// ---- DUTs/ST_MoverStatus.TcDUT
// C# 端對應 MoverStatus (Pack = 1)
{attribute 'pack_mode' := '1'}
TYPE ST_MoverStatus :
STRUCT
    fPositionMm : LREAL;    // 環上位置 (mm), 0~3000
    fVelocityMmS : LREAL;   // 實際速度 (mm/s)
    bPowered : BOOL;
    bBusy : BOOL;
    bDone : BOOL;
    bError : BOOL;
    nErrorId : UDINT;
    bHasPart : BOOL;        // 有工件
    bPressed : BOOL;        // 已下壓
    nStation : INT;         // 停在哪一站，0 = 不在站上
END_STRUCT
END_TYPE

// ---- DUTs/ST_StationStatus.TcDUT
// C# 端對應 StationStatus (Pack = 1)
{attribute 'pack_mode' := '1'}
TYPE ST_StationStatus :
STRUCT
    eState : E_StationState;
    nStep : INT;            // 站內步驟，見 README
    bOccupied : BOOL;       // 站內有 mover 或站在動作
    nMover : INT;           // 處理中的 mover，0 = 無
    bError : BOOL;
    nErrorId : UDINT;
    nDoneCount : UDINT;     // 完成次數
    fAxis1Mm : LREAL;       // X (mm)；下壓站不用
    fAxis2Mm : LREAL;       // Y (mm)；下壓站不用
    fAxis3Mm : LREAL;       // Z (mm)，往下為正
    bGripClosed : BOOL;     // 夾爪閉合；下壓站固定 FALSE
END_STRUCT
END_TYPE

// ---- GVLs/GVL_ErrorId.TcGVL
// 應用程式錯誤碼；MC / NC 的錯誤碼照原值傳出
{attribute 'qualified_only'}
VAR_GLOBAL CONSTANT
    cErrInvalidState : UDINT := 16#E001;        // 狀態機進到未定義狀態
    cErrMoveTimeout : UDINT := 16#E101;         // mover 移動逾時
    cErrStationTimeout : UDINT := 16#E201;      // 站內步驟逾時
    cErrInitTimeout : UDINT := 16#E301;         // 初始化步驟逾時
    cErrEnvInit : UDINT := 16#E302;             // Utility 環境 Init 失敗
    cErrIdDetection : UDINT := 16#E303;         // Mover ID detection 失敗
    cErrGroup : UDINT := 16#E304;               // CA group enable 失敗
    cErrLostReady : UDINT := 16#E310;           // 執行中掉出可控
    cErrCycle : UDINT := 16#E401;               // 自動循環失敗
END_VAR

// ---- GVLs/GVL_Param.TcGVL
{attribute 'qualified_only'}
VAR_GLOBAL CONSTANT
    cMoverCount : INT := 4;                     // mover 數，與 XTS 設定一致
    cStationCount : INT := 3;                   // 站數
    cStationLoad : INT := 1;                    // 站號：Load
    cStationPress : INT := 2;                   // 站號：Press
    cStationUnload : INT := 3;                  // 站號：Unload
    cTrackLengthMm : LREAL := 3000.0;           // 軌道長 (mm)
    cStationPosMm : ARRAY[1..3] OF LREAL := [1600.0, 2100.0, 2600.0];   // 各站 mover 停止位置 (mm, 環上)
    cMaxVelocityMmS : LREAL := 1500.0;          // mover 速度上限 (mm/s)
    cDefaultVelocityMmS : LREAL := 400.0;       // 自動循環 / 送站速度 (mm/s)
    cMoverAccMmS2 : LREAL := 2000.0;            // mover 加減速度 (mm/s2)
    cMoverJerkMmS3 : LREAL := 20000.0;          // mover jerk (mm/s3)
    cCaGapMm : LREAL := 110.0;                  // CA 最小間距 (mm)
    cAtStationTolMm : LREAL := 1.0;             // 判定到站的容差 (mm)
    cMoveTimeout : TIME := T#10M;               // mover 單次移動上限
    cInitStepTimeout : TIME := T#5M;            // 初始化每一步上限，UmRT 偏慢所以放寬
    cResetTime : TIME := T#500MS;               // 初始化 reset 保持時間
    cStationStepTimeout : TIME := T#2M;         // 站內每一步上限
    cGantryAxisCount : INT := 3;                // XYZ 軸數
    cAxisX : INT := 1;
    cAxisY : INT := 2;
    cAxisZ : INT := 3;
    cGantryVelocityMmS : LREAL := 200.0;        // XYZ 與下壓軸速度 (mm/s)
    cGantryAccMmS2 : LREAL := 1000.0;           // XYZ 與下壓軸加減速度 (mm/s2)
    cGantryZUpMm : LREAL := 0.0;                // Z 上位 (mm)
    cGantryZDownMm : LREAL := 80.0;             // Z 下位 (mm)
    cGantryFeederXMm : LREAL := 300.0;          // Load 取料點 X (mm)
    cGantryFeederYMm : LREAL := 150.0;          // Load 取料點 Y (mm)
    cGantryOutXMm : LREAL := 300.0;             // Unload 放料點 X (mm)
    cGantryOutYMm : LREAL := -150.0;            // Unload 放料點 Y (mm)
    cGantryMoverXMm : LREAL := 0.0;             // mover 正上方 X (mm)
    cGantryMoverYMm : LREAL := 0.0;             // mover 正上方 Y (mm)
    cGripTime : TIME := T#300MS;                // 夾 / 放 時間
    cPressZDownMm : LREAL := 50.0;              // 下壓位置 (mm)
    cPressHoldTime : TIME := T#1S;              // 保壓時間
END_VAR

// ---- POUs/MAIN.TcPOU
PROGRAM MAIN
VAR
    aAxis : ARRAY[1..GVL_Param.cMoverCount] OF AXIS_REF;              // 連 NC Mover Axis 1..4
    stCaGroup : Tc3_McCoordinatedMotion.AXES_GROUP_REF;                 // 連 XtsCaGroup
    aLoadAxis : ARRAY[1..GVL_Param.cGantryAxisCount] OF AXIS_REF;      // 連 Load X / Y / Z
    aUnloadAxis : ARRAY[1..GVL_Param.cGantryAxisCount] OF AXIS_REF;    // 連 Unload X / Y / Z
    stPressAxis : AXIS_REF;                                             // 連 Press Z
    fbXts : FB_XTS_Control;                                             // C# RPC 主入口：MAIN.fbXts
    refMover1 : REFERENCE TO FB_Mover;                                  // 備案 RPC 路徑：MAIN.refMover1..4
    refMover2 : REFERENCE TO FB_Mover;
    refMover3 : REFERENCE TO FB_Mover;
    refMover4 : REFERENCE TO FB_Mover;
END_VAR

fbXts(aMoverAxis := aAxis, stGroup := stCaGroup, aLoadAxis := aLoadAxis,
    aUnloadAxis := aUnloadAxis, stPressAxis := stPressAxis);
// REFERENCE 每 cycle 重取 (PTR-03)
refMover1 REF= fbXts.M_GetMover(1);
refMover2 REF= fbXts.M_GetMover(2);
refMover3 REF= fbXts.M_GetMover(3);
refMover4 REF= fbXts.M_GetMover(4);

END_PROGRAM

// ---- POUs/FB_XTS_Control.TcPOU
// 整線總控：初始化 (Find mover 1 → 送電 → CA group)、模式、自動循環 Load → Press → Unload、派 mover 到站。
// 擁有 4 個 FB_Mover 與 3 個站；每 cycle 把 ST_CmdPermit 寫給子 FB，所有命令檢查只走 F_CheckCmdAllowed。
FUNCTION_BLOCK FB_XTS_Control
VAR_IN_OUT
    aMoverAxis : ARRAY[1..GVL_Param.cMoverCount] OF AXIS_REF;          // XTS mover NC 軸
    stGroup : Tc3_McCoordinatedMotion.AXES_GROUP_REF;                   // CA group
    aLoadAxis : ARRAY[1..GVL_Param.cGantryAxisCount] OF AXIS_REF;      // Load 站 XYZ
    aUnloadAxis : ARRAY[1..GVL_Param.cGantryAxisCount] OF AXIS_REF;    // Unload 站 XYZ
    stPressAxis : AXIS_REF;                                             // Press 站下壓軸
END_VAR
VAR_OUTPUT
    bReady : BOOL;                  // 可控
    eMode : E_XtsMode;
    eInitStep : E_InitStep;
    eCycleState : E_CycleState;
    bError : BOOL;
    nErrorId : UDINT;
END_VAR
VAR
    aMover : ARRAY[1..GVL_Param.cMoverCount] OF FB_Mover;
    fbLoad : FB_StationLoad;
    fbPress : FB_StationPress;
    fbUnload : FB_StationUnload;
    aStationPtr : ARRAY[1..GVL_Param.cStationCount] OF POINTER TO FB_Station;   // 每 cycle 重取
    fbEnvironment : Tc3_XTS_Utility.FB_TcIoXtsEnvironment;
    stEnvConfig : Tc3_XTS_Utility.ST_XtsEnvironmentConfiguration;
    fbGroup : FB_CaGroup;
    fbInitTimer : TON;
    fbResetTimer : TON;
    stPermit : ST_CmdPermit;
    stStatus : ST_LineStatus;       // M_GetStatus 回傳的快照
    sInitMsg : STRING;              // 初始化進度或失敗原因
    sCycleMsg : STRING;             // 自動循環訊息
    bEnvInitialized : BOOL;
    bPowerOn : BOOL;
    bGroupEnable : BOOL;
    bInitReset : BOOL;
    eInitStepLast : E_InitStep;
    tInitStart : TIME;              // M_InitialXTS 被取走的時刻
    nFindMover1Ms : UDINT;          // 各步完成時間 (ms，從 tInitStart 起算；0 = 這次還沒完成)
    bFindMover1Detected : BOOL;     // TRUE = detection valid；FALSE 且 nFindMover1Ms > 0 = 跳過
    nPowerOnMs : UDINT;
    nGroupMs : UDINT;
    bReqInit : BOOL;                // method 設，body 取走
    bReqStop : BOOL;
    bReqSetMode : BOOL;
    eReqMode : E_XtsMode;
    bReqStartCycle : BOOL;
    nReqCycleMover : INT;
    bStopPulse : BOOL;              // 本 cycle 對站送 abort
    nCycleMover : INT;
    nCycleStation : INT;
    bCycleMoveIssued : BOOL;
    nCycleCount : UDINT;
    tCycleStart : TIME;
    aStationDoneMs : ARRAY[1..GVL_Param.cStationCount] OF UDINT;
    aLastDoneCount : ARRAY[1..GVL_Param.cStationCount] OF UDINT;
    aMoverAtStation : ARRAY[1..GVL_Param.cStationCount] OF INT;
    pStation : POINTER TO FB_Station;
    bAllPowered : BOOL;
    bAnyMoverError : BOOL;
    bInitBusy : BOOL;
    fDistMm : LREAL;
    i : INT;
    j : INT;
    nStation : INT;
END_VAR

// 1. 站指標每 cycle 重取 (PTR-03)
aStationPtr[GVL_Param.cStationLoad] := ADR(fbLoad);
aStationPtr[GVL_Param.cStationPress] := ADR(fbPress);
aStationPtr[GVL_Param.cStationUnload] := ADR(fbUnload);

// 2. 取走 method 設的命令
bStopPulse := FALSE;
IF bReqStop THEN
    bReqStop := FALSE;
    bStopPulse := TRUE;
    FOR i := 1 TO GVL_Param.cMoverCount DO
        aMover[i].M_Stop();
    END_FOR
    IF (eCycleState = E_CycleState.ToStation) OR (eCycleState = E_CycleState.InStation) THEN
        eCycleState := E_CycleState.Stopped;
        sCycleMsg := 'Stopped by M_Stop';
    END_IF
END_IF
IF bReqSetMode THEN
    bReqSetMode := FALSE;
    eMode := eReqMode;
END_IF
IF bReqInit THEN
    bReqInit := FALSE;
    bError := FALSE;
    nErrorId := 0;
    sInitMsg := 'Reset';
    eInitStep := E_InitStep.Reset;
    tInitStart := TIME();
    nFindMover1Ms := 0;
    bFindMover1Detected := FALSE;
    nPowerOnMs := 0;
    nGroupMs := 0;
END_IF

// 3. 初始化：Find mover 1 → 送電 → CA group
bInitBusy := M_InitBusy();
fbInitTimer(IN := bInitBusy AND (eInitStep = eInitStepLast), PT := GVL_Param.cInitStepTimeout);
eInitStepLast := eInitStep;
fbResetTimer(IN := (eInitStep = E_InitStep.Reset), PT := GVL_Param.cResetTime);
CASE eInitStep OF
E_InitStep.Idle, E_InitStep.Ready, E_InitStep.Error:
    ;
E_InitStep.Reset:
    bInitReset := TRUE;
    bPowerOn := FALSE;
    bGroupEnable := FALSE;
    IF fbResetTimer.Q THEN
        bInitReset := FALSE;
        IF bEnvInitialized THEN
            eInitStep := E_InitStep.WaitMovers;
        ELSE
            stEnvConfig.bEnableInitInfoServer := TRUE;
            stEnvConfig.bEnableInitCaGroup := TRUE;
            fbEnvironment.P_XtsEnvironmentConfiguration := stEnvConfig;
            eInitStep := E_InitStep.InitEnvironment;
        END_IF
        sInitMsg := F_InitStepName(eInitStep);
    END_IF
E_InitStep.InitEnvironment:
    // Init 是非同步的，回 TRUE 才算做完
    IF fbEnvironment.Init(TRUE) THEN
        fbEnvironment.Init(FALSE);
        IF fbEnvironment.P_IsInitialized THEN
            bEnvInitialized := TRUE;
            eInitStep := E_InitStep.WaitMovers;
            sInitMsg := F_InitStepName(eInitStep);
        ELSE
            M_SetInitError(nId := GVL_ErrorId.cErrEnvInit, sText := 'Tc3_XTS_Utility Init failed');
        END_IF
    END_IF
E_InitStep.WaitMovers:
    IF (fbEnvironment.XpuTcIo(1).GetDetectedMoverCount() = INT_TO_UDINT(GVL_Param.cMoverCount))
        AND fbEnvironment.XpuTcIo(1).GetAreAllPositionsValid() THEN
        eInitStep := E_InitStep.FindMover1;
        sInitMsg := F_InitStepName(eInitStep);
    END_IF
E_InitStep.FindMover1:
    // 專案設定 IdDetectionMode = Mover1；detection 要在 MC_Power 之前 (XTS 事件 9016)
    IF fbEnvironment.XpuTcIo(1).GetMoverIdDetectionMode() = MoverIdDetectionMode.Mover1 THEN
        IF fbEnvironment.XpuTcIo(1).TriggerMoverIdDetection() THEN
            eInitStep := E_InitStep.FindMover1Wait;
            sInitMsg := 'FindMover1: Mover ID detection triggered, waiting for result';
        ELSE
            M_SetInitError(nId := GVL_ErrorId.cErrIdDetection, sText := 'TriggerMoverIdDetection rejected');
        END_IF
    ELSE
        // 防呆：XPU 被改回 Standard 時不做 detection，mover 編號照設定順序
        eInitStep := E_InitStep.PowerOn;
        sInitMsg := 'FindMover1 skipped: XPU IdDetectionMode is not Mover1, PowerOn';
        nFindMover1Ms := MAX(TIME_TO_UDINT(TIME() - tInitStart), 1);
    END_IF
E_InitStep.FindMover1Wait:
    IF fbEnvironment.XpuTcIo(1).GetHasMoverIdDetectionError() THEN
        M_SetInitError(nId := GVL_ErrorId.cErrIdDetection, sText := 'Mover ID detection error');
    ELSIF fbEnvironment.XpuTcIo(1).GetIsMoverIdDetectionValid() THEN
        eInitStep := E_InitStep.PowerOn;
        sInitMsg := 'FindMover1 done (Mover ID detection valid), PowerOn';
        nFindMover1Ms := MAX(TIME_TO_UDINT(TIME() - tInitStart), 1);
        bFindMover1Detected := TRUE;
    END_IF
E_InitStep.PowerOn:
    bPowerOn := TRUE;
    IF bAllPowered AND fbLoad.bAxesPowered AND fbPress.bAxesPowered AND fbUnload.bAxesPowered THEN
        eInitStep := E_InitStep.EnableGroup;
        sInitMsg := F_InitStepName(eInitStep);
        nPowerOnMs := MAX(TIME_TO_UDINT(TIME() - tInitStart), 1);
    END_IF
E_InitStep.EnableGroup:
    bGroupEnable := TRUE;
    IF fbGroup.bError THEN
        M_SetInitError(nId := fbGroup.nErrorId, sText := 'CA group error');
    ELSIF fbGroup.bReady THEN
        eInitStep := E_InitStep.Ready;
        sInitMsg := 'Ready';
        nGroupMs := MAX(TIME_TO_UDINT(TIME() - tInitStart), 1);
    END_IF
ELSE
    M_SetInitError(nId := GVL_ErrorId.cErrInvalidState, sText := 'invalid init step');
END_CASE
IF fbInitTimer.Q THEN
    M_SetInitError(nId := GVL_ErrorId.cErrInitTimeout, sText := 'step timeout');
END_IF

// 4. 可控監視：任何 mover error、失電、group 失效、站上軸 error 都掉出 ready
bAllPowered := TRUE;
bAnyMoverError := FALSE;
FOR i := 1 TO GVL_Param.cMoverCount DO
    bAllPowered := bAllPowered AND aMover[i].bPowered;
    bAnyMoverError := bAnyMoverError OR aMover[i].bError;
END_FOR
IF eInitStep = E_InitStep.Ready THEN
    IF bAnyMoverError THEN
        M_SetInitError(nId := GVL_ErrorId.cErrLostReady, sText := 'mover error');
    ELSIF NOT bAllPowered THEN
        M_SetInitError(nId := GVL_ErrorId.cErrLostReady, sText := 'mover power lost');
    ELSIF NOT fbGroup.bReady THEN
        M_SetInitError(nId := GVL_ErrorId.cErrLostReady, sText := 'CA group not ready');
    ELSIF fbLoad.bAxisError OR fbPress.bAxisError OR fbUnload.bAxisError THEN
        M_SetInitError(nId := GVL_ErrorId.cErrLostReady, sText := 'station axis error');
    END_IF
END_IF
bReady := (eInitStep = E_InitStep.Ready);
stPermit.bReady := bReady;
stPermit.eMode := eMode;

// 5. 哪個 mover 停在哪一站 (停止且在容差內)
FOR nStation := 1 TO GVL_Param.cStationCount DO
    aMoverAtStation[nStation] := 0;
    FOR i := 1 TO GVL_Param.cMoverCount DO
        fDistMm := F_RingPosition(fPositionMm := aMover[i].fPositionMm - GVL_Param.cStationPosMm[nStation]
            + GVL_Param.cTrackLengthMm / 2.0, fLengthMm := GVL_Param.cTrackLengthMm) - GVL_Param.cTrackLengthMm / 2.0;
        IF NOT aMover[i].bBusy AND (ABS(fDistMm) <= GVL_Param.cAtStationTolMm) THEN
            aMoverAtStation[nStation] := i;
        END_IF
    END_FOR
    pStation := aStationPtr[nStation];
    IF pStation <> 0 THEN
        pStation^.nMoverAtStation := aMoverAtStation[nStation];
        j := aMoverAtStation[nStation];
        IF j > 0 THEN
            pStation^.bMoverHasPart := aMover[j].bHasPart;
            pStation^.bMoverPressed := aMover[j].bPressed;
        ELSE
            pStation^.bMoverHasPart := FALSE;
            pStation^.bMoverPressed := FALSE;
        END_IF
    END_IF
END_FOR

// 6. 站完成 → 更新 mover 工件狀態 (手動與自動都走這裡)
FOR nStation := 1 TO GVL_Param.cStationCount DO
    pStation := aStationPtr[nStation];
    IF pStation <> 0 THEN
        IF pStation^.nDoneCount <> aLastDoneCount[nStation] THEN
            aLastDoneCount[nStation] := pStation^.nDoneCount;
            j := pStation^.nMover;
            IF (j >= 1) AND (j <= GVL_Param.cMoverCount) THEN
                CASE nStation OF
                GVL_Param.cStationLoad:
                    aMover[j].M_SetPart(bPart := TRUE, bPress := FALSE);
                GVL_Param.cStationPress:
                    aMover[j].M_SetPart(bPart := aMover[j].bHasPart, bPress := TRUE);
                GVL_Param.cStationUnload:
                    aMover[j].M_SetPart(bPart := FALSE, bPress := FALSE);
                END_CASE
            END_IF
        END_IF
    END_IF
END_FOR

// 7. 自動循環：mover 依序到 Load → Press → Unload
IF NOT bReady AND ((eCycleState = E_CycleState.ToStation) OR (eCycleState = E_CycleState.InStation)) THEN
    eCycleState := E_CycleState.Error;
    sCycleMsg := 'Lost ready during cycle';
END_IF
pStation := 0;
IF (nCycleStation >= 1) AND (nCycleStation <= GVL_Param.cStationCount) THEN
    pStation := aStationPtr[nCycleStation];
END_IF
CASE eCycleState OF
E_CycleState.Idle, E_CycleState.Done, E_CycleState.Stopped, E_CycleState.Error:
    IF bReqStartCycle THEN
        nCycleMover := nReqCycleMover;
        nCycleStation := GVL_Param.cStationLoad;
        bCycleMoveIssued := FALSE;
        tCycleStart := TIME();
        FOR nStation := 1 TO GVL_Param.cStationCount DO
            aStationDoneMs[nStation] := 0;
        END_FOR
        sCycleMsg := 'Cycle started';
        eCycleState := E_CycleState.ToStation;
    END_IF
E_CycleState.ToStation:
    IF pStation = 0 THEN
        eCycleState := E_CycleState.Error;
        sCycleMsg := 'Invalid station index';
    ELSIF NOT bCycleMoveIssued THEN
        bCycleMoveIssued := aMover[nCycleMover].M_RequestMove(fPosition := GVL_Param.cStationPosMm[nCycleStation],
            fVelocity := GVL_Param.cDefaultVelocityMmS, sMsg => sCycleMsg);
    ELSIF aMover[nCycleMover].bDone AND (aMoverAtStation[nCycleStation] = nCycleMover) THEN
        IF pStation^.M_RequestStart(sMsg => sCycleMsg) THEN
            eCycleState := E_CycleState.InStation;
        ELSE
            eCycleState := E_CycleState.Error;
        END_IF
    END_IF
E_CycleState.InStation:
    IF pStation = 0 THEN
        eCycleState := E_CycleState.Error;
        sCycleMsg := 'Invalid station index';
    ELSIF pStation^.eState = E_StationState.Error THEN
        eCycleState := E_CycleState.Error;
        sCycleMsg := 'Station error';
    ELSIF pStation^.eState = E_StationState.Done THEN
        aStationDoneMs[nCycleStation] := TIME_TO_UDINT(TIME() - tCycleStart);
        pStation^.M_RequestRelease(sMsg => sCycleMsg);
        IF nCycleStation < GVL_Param.cStationCount THEN
            nCycleStation := nCycleStation + 1;
            bCycleMoveIssued := FALSE;
            eCycleState := E_CycleState.ToStation;
        ELSE
            nCycleCount := nCycleCount + 1;
            sCycleMsg := 'Cycle done';
            eCycleState := E_CycleState.Done;
        END_IF
    END_IF
ELSE
    eCycleState := E_CycleState.Error;
    sCycleMsg := 'Invalid cycle state';
END_CASE
bReqStartCycle := FALSE;

// 8. 呼叫子 FB (每 cycle 無條件)
FOR i := 1 TO GVL_Param.cMoverCount DO
    aMover[i](nIndex := i, stPermit := stPermit, bPowerEnable := bPowerOn, bResetCmd := bInitReset,
        stAxis := aMoverAxis[i]);
END_FOR
fbGroup(Group := stGroup, Axes := aMoverAxis, bEnable := bGroupEnable, bReset := bInitReset);
fbLoad(nIndex := GVL_Param.cStationLoad, stPermit := stPermit, bPowerEnable := bPowerOn,
    bResetCmd := bInitReset, bAbort := bStopPulse, aAxis := aLoadAxis);
fbPress(nIndex := GVL_Param.cStationPress, stPermit := stPermit, bPowerEnable := bPowerOn,
    bResetCmd := bInitReset, bAbort := bStopPulse, stAxis := stPressAxis);
fbUnload(nIndex := GVL_Param.cStationUnload, stPermit := stPermit, bPowerEnable := bPowerOn,
    bResetCmd := bInitReset, bAbort := bStopPulse, aAxis := aUnloadAxis);

// 9. 狀態快照
stStatus.bReady := bReady;
stStatus.eMode := eMode;
stStatus.eInitStep := eInitStep;
stStatus.bError := bError;
stStatus.nErrorId := nErrorId;
stStatus.eCycleState := eCycleState;
stStatus.nCycleMover := nCycleMover;
stStatus.nCycleStation := nCycleStation;
stStatus.nCycleCount := nCycleCount;
FOR i := 1 TO GVL_Param.cMoverCount DO
    stStatus.aMover[i].fPositionMm := aMover[i].fPositionMm;
    stStatus.aMover[i].fVelocityMmS := aMover[i].fVelocityMmS;
    stStatus.aMover[i].bPowered := aMover[i].bPowered;
    stStatus.aMover[i].bBusy := aMover[i].bBusy;
    stStatus.aMover[i].bDone := aMover[i].bDone;
    stStatus.aMover[i].bError := aMover[i].bError;
    stStatus.aMover[i].nErrorId := aMover[i].nErrorId;
    stStatus.aMover[i].bHasPart := aMover[i].bHasPart;
    stStatus.aMover[i].bPressed := aMover[i].bPressed;
    stStatus.aMover[i].nStation := 0;
END_FOR
FOR nStation := 1 TO GVL_Param.cStationCount DO
    stStatus.aStationDoneMs[nStation] := aStationDoneMs[nStation];
    j := aMoverAtStation[nStation];
    IF (j >= 1) AND (j <= GVL_Param.cMoverCount) THEN
        stStatus.aMover[j].nStation := nStation;
    END_IF
    pStation := aStationPtr[nStation];
    IF pStation <> 0 THEN
        stStatus.aStation[nStation] := pStation^.M_GetStatusStruct();
    END_IF
END_FOR

// 內部用：給 MAIN 的 REFERENCE 備案路徑。超出範圍回 mover 1。
METHOD PUBLIC M_GetMover : REFERENCE TO FB_Mover
VAR_INPUT
    nMover : INT;
END_VAR
M_GetMover REF= aMover[LIMIT(1, nMover, GVL_Param.cMoverCount)];
END_METHOD

// RPC：整線快照 (mover、站、XYZ / 下壓軸位置、循環)，隨時可讀
{attribute 'TcRpcEnable'}
METHOD PUBLIC M_GetStatus : BOOL
VAR_OUTPUT
    stLine : ST_LineStatus;
    sCycle : STRING;            // 自動循環訊息
END_VAR
stLine := stStatus;
sCycle := sCycleMsg;
M_GetStatus := TRUE;
END_METHOD

METHOD PRIVATE M_InitBusy : BOOL
M_InitBusy := (eInitStep = E_InitStep.Reset) OR (eInitStep = E_InitStep.InitEnvironment)
    OR (eInitStep = E_InitStep.WaitMovers) OR (eInitStep = E_InitStep.FindMover1)
    OR (eInitStep = E_InitStep.FindMover1Wait) OR (eInitStep = E_InitStep.PowerOn)
    OR (eInitStep = E_InitStep.EnableGroup);
END_METHOD

// RPC：開始初始化 (Reset → Find mover 1 → PowerOn → EnableGroup)。回 TRUE = 已接受，用 M_ReadXTS_Status 看進度。
{attribute 'TcRpcEnable'}
METHOD PUBLIC M_InitialXTS : BOOL
VAR_OUTPUT
    sMsg : STRING;
END_VAR
M_InitialXTS := FALSE;
IF bReqInit THEN
    sMsg := 'Previous command not yet taken by PLC, retry';
ELSIF M_InitBusy() THEN
    sMsg := CONCAT('Init already running: ', F_InitStepName(eInitStep));
ELSIF (eCycleState = E_CycleState.ToStation) OR (eCycleState = E_CycleState.InStation) THEN
    sMsg := 'Cycle running, call M_Stop first';
ELSIF bReady THEN
    sMsg := 'Already ready';
ELSE
    bReqInit := TRUE;
    sMsg := 'Init started';
    M_InitialXTS := TRUE;
END_IF
END_METHOD

// RPC：總控層的 mover 移動 (陣列元素路徑不能用時的備案)。需 ready + Manual。
{attribute 'TcRpcEnable'}
METHOD PUBLIC M_MoveTo : BOOL
VAR_INPUT
    nMover : UINT;              // 1..cMoverCount
    fPosition : LREAL;          // 目標環上位置 (mm)
    fVelocity : LREAL;          // 速度 (mm/s)
END_VAR
VAR_OUTPUT
    sMsg : STRING;
END_VAR
M_MoveTo := FALSE;
IF NOT F_CheckCmdAllowed(stPermit := stPermit, bNeedManual := TRUE, bNeedAuto := FALSE, sMsg => sMsg) THEN
    RETURN;
END_IF
IF (nMover < 1) OR (nMover > INT_TO_UINT(GVL_Param.cMoverCount)) THEN
    sMsg := CONCAT('nMover out of range 1..', INT_TO_STRING(GVL_Param.cMoverCount));
    RETURN;
END_IF
M_MoveTo := aMover[UINT_TO_INT(nMover)].M_RequestMove(fPosition := fPosition, fVelocity := fVelocity, sMsg => sMsg);
END_METHOD

// RPC：可控閘門狀態，隨時可讀
{attribute 'TcRpcEnable'}
METHOD PUBLIC M_ReadXTS_Status : BOOL
VAR_OUTPUT
    bIsReady : BOOL;            // TRUE 才能下站與 mover 命令
    eStep : E_InitStep;         // 初始化目前步驟
    sStepMsg : STRING;          // 進度或失敗原因
    bIsError : BOOL;
    nErrId : UDINT;
    eModeNow : E_XtsMode;
    nFindMover1DoneMs : UDINT;  // 各步完成時間 (PLC ms，從 M_InitialXTS 被取走起算；0 = 這次還沒完成)
    bFindMover1Valid : BOOL;    // TRUE = Mover ID detection valid；FALSE 且時間 > 0 = IdDetectionMode 不是 Mover1、跳過
    nPowerOnDoneMs : UDINT;
    nGroupDoneMs : UDINT;
END_VAR
bIsReady := bReady;
eStep := eInitStep;
sStepMsg := sInitMsg;
bIsError := bError;
nErrId := nErrorId;
eModeNow := eMode;
nFindMover1DoneMs := nFindMover1Ms;
bFindMover1Valid := bFindMover1Detected;
nPowerOnDoneMs := nPowerOnMs;
nGroupDoneMs := nGroupMs;
M_ReadXTS_Status := TRUE;
END_METHOD

// RPC：總控層的手動放行 (備案路徑)。需 ready + Manual。
{attribute 'TcRpcEnable'}
METHOD PUBLIC M_ReleaseStation : BOOL
VAR_INPUT
    nStation : UINT;            // 1 = Load, 2 = Press, 3 = Unload
END_VAR
VAR_OUTPUT
    sMsg : STRING;
END_VAR
VAR
    pSt : POINTER TO FB_Station;
END_VAR
M_ReleaseStation := FALSE;
IF NOT F_CheckCmdAllowed(stPermit := stPermit, bNeedManual := TRUE, bNeedAuto := FALSE, sMsg => sMsg) THEN
    RETURN;
END_IF
IF (nStation < 1) OR (nStation > INT_TO_UINT(GVL_Param.cStationCount)) THEN
    sMsg := CONCAT('nStation out of range 1..', INT_TO_STRING(GVL_Param.cStationCount));
    RETURN;
END_IF
pSt := aStationPtr[UINT_TO_INT(nStation)];
IF pSt = 0 THEN
    sMsg := 'Station not ready yet, retry';
    RETURN;
END_IF
M_ReleaseStation := pSt^.M_RequestRelease(sMsg => sMsg);
END_METHOD

// RPC：把 mover 送到指定站。需 ready + Manual、站號有效、站沒被其他 mover 佔用。
{attribute 'TcRpcEnable'}
METHOD PUBLIC M_SendToStation : BOOL
VAR_INPUT
    nMover : UINT;              // 1..cMoverCount
    nStation : UINT;            // 1 = Load, 2 = Press, 3 = Unload
END_VAR
VAR_OUTPUT
    sMsg : STRING;
END_VAR
VAR
    nMv : INT;
    nSt : INT;
END_VAR
M_SendToStation := FALSE;
IF NOT F_CheckCmdAllowed(stPermit := stPermit, bNeedManual := TRUE, bNeedAuto := FALSE, sMsg => sMsg) THEN
    RETURN;
END_IF
IF (nMover < 1) OR (nMover > INT_TO_UINT(GVL_Param.cMoverCount)) THEN
    sMsg := CONCAT('nMover out of range 1..', INT_TO_STRING(GVL_Param.cMoverCount));
    RETURN;
END_IF
IF (nStation < 1) OR (nStation > INT_TO_UINT(GVL_Param.cStationCount)) THEN
    sMsg := CONCAT('nStation out of range 1..', INT_TO_STRING(GVL_Param.cStationCount));
    RETURN;
END_IF
nMv := UINT_TO_INT(nMover);       // 已檢查範圍，不會溢位
nSt := UINT_TO_INT(nStation);
IF (aMoverAtStation[nSt] <> 0) AND (aMoverAtStation[nSt] <> nMv) THEN
    sMsg := CONCAT(CONCAT('Station occupied by mover ', INT_TO_STRING(aMoverAtStation[nSt])), ', move it away first');
    RETURN;
END_IF
M_SendToStation := aMover[nMv].M_RequestMove(fPosition := GVL_Param.cStationPosMm[nSt],
    fVelocity := GVL_Param.cDefaultVelocityMmS, sMsg => sMsg);
END_METHOD

METHOD PRIVATE M_SetInitError
VAR_INPUT
    nId : UDINT;
    sText : STRING;
END_VAR
sInitMsg := CONCAT(CONCAT(F_InitStepName(eInitStep), ': '), sText);
bError := TRUE;
nErrorId := nId;
IF nErrorId = 0 THEN
    nErrorId := GVL_ErrorId.cErrInvalidState;
END_IF
eInitStep := E_InitStep.Error;
END_METHOD

// RPC：切換模式 0 = Manual、1 = Auto。自動循環中拒絕。不受 ready 限制。
{attribute 'TcRpcEnable'}
METHOD PUBLIC M_SetMode : BOOL
VAR_INPUT
    nMode : INT;                // 0 = Manual, 1 = Auto
END_VAR
VAR_OUTPUT
    sMsg : STRING;
END_VAR
M_SetMode := FALSE;
IF (eCycleState = E_CycleState.ToStation) OR (eCycleState = E_CycleState.InStation) THEN
    sMsg := 'Cycle running, call M_Stop first';
ELSIF nMode = 0 THEN
    eReqMode := E_XtsMode.Manual;
    bReqSetMode := TRUE;
    sMsg := 'Mode -> Manual';
    M_SetMode := TRUE;
ELSIF nMode = 1 THEN
    eReqMode := E_XtsMode.Auto;
    bReqSetMode := TRUE;
    sMsg := 'Mode -> Auto';
    M_SetMode := TRUE;
ELSE
    sMsg := 'nMode must be 0 (Manual) or 1 (Auto)';
END_IF
END_METHOD

// RPC：nMover 跑一輪 Load → Press → Unload。需 ready + Auto、三站 Idle、mover 沒工件、路徑上沒有其他 mover。
{attribute 'TcRpcEnable'}
METHOD PUBLIC M_StartCycle : BOOL
VAR_INPUT
    nMover : UINT;              // 1..cMoverCount
END_VAR
VAR_OUTPUT
    sMsg : STRING;
END_VAR
VAR
    nMv : INT;
    nOther : INT;
    fPathMm : LREAL;            // 到 Unload 的路徑長 + CA 間距 (mm)
    fAheadMm : LREAL;           // 其他 mover 在前方多遠 (mm)
END_VAR
M_StartCycle := FALSE;
IF NOT F_CheckCmdAllowed(stPermit := stPermit, bNeedManual := FALSE, bNeedAuto := TRUE, sMsg => sMsg) THEN
    RETURN;
END_IF
IF bReqStartCycle THEN
    sMsg := 'Previous command not yet taken by PLC, retry';
    RETURN;
END_IF
IF (eCycleState = E_CycleState.ToStation) OR (eCycleState = E_CycleState.InStation) THEN
    sMsg := 'Cycle already running';
    RETURN;
END_IF
IF (nMover < 1) OR (nMover > INT_TO_UINT(GVL_Param.cMoverCount)) THEN
    sMsg := CONCAT('nMover out of range 1..', INT_TO_STRING(GVL_Param.cMoverCount));
    RETURN;
END_IF
nMv := UINT_TO_INT(nMover);       // 已檢查範圍，不會溢位
IF aMover[nMv].bHasPart THEN
    sMsg := 'Mover already has a part, unload it first';
    RETURN;
END_IF
IF aMover[nMv].bBusy OR aMover[nMv].bError THEN
    sMsg := 'Mover busy or in error';
    RETURN;
END_IF
IF (fbLoad.eState <> E_StationState.Idle) OR (fbPress.eState <> E_StationState.Idle)
    OR (fbUnload.eState <> E_StationState.Idle) THEN
    sMsg := 'All stations must be Idle';
    RETURN;
END_IF
// CA 會讓 mover 排在前車後面，路徑上有車就到不了站
fPathMm := F_RingPosition(fPositionMm := GVL_Param.cStationPosMm[GVL_Param.cStationUnload] - aMover[nMv].fPositionMm,
    fLengthMm := GVL_Param.cTrackLengthMm) + GVL_Param.cCaGapMm;
FOR nOther := 1 TO GVL_Param.cMoverCount DO
    IF nOther <> nMv THEN
        fAheadMm := F_RingPosition(fPositionMm := aMover[nOther].fPositionMm - aMover[nMv].fPositionMm,
            fLengthMm := GVL_Param.cTrackLengthMm);
        IF fAheadMm < fPathMm THEN
            sMsg := CONCAT(CONCAT('Mover ', INT_TO_STRING(nOther)), ' is in the path, move it away in Manual first');
            RETURN;
        END_IF
    END_IF
END_FOR
nReqCycleMover := nMv;
bReqStartCycle := TRUE;
sMsg := 'Cycle accepted';
M_StartCycle := TRUE;
END_METHOD

// RPC：總控層的手動站啟動 (子類別上繼承來的 RPC 不能用時的備案)。需 ready + Manual。
{attribute 'TcRpcEnable'}
METHOD PUBLIC M_StartStation : BOOL
VAR_INPUT
    nStation : UINT;            // 1 = Load, 2 = Press, 3 = Unload
END_VAR
VAR_OUTPUT
    sMsg : STRING;
END_VAR
VAR
    pSt : POINTER TO FB_Station;
END_VAR
M_StartStation := FALSE;
IF NOT F_CheckCmdAllowed(stPermit := stPermit, bNeedManual := TRUE, bNeedAuto := FALSE, sMsg => sMsg) THEN
    RETURN;
END_IF
IF (nStation < 1) OR (nStation > INT_TO_UINT(GVL_Param.cStationCount)) THEN
    sMsg := CONCAT('nStation out of range 1..', INT_TO_STRING(GVL_Param.cStationCount));
    RETURN;
END_IF
pSt := aStationPtr[UINT_TO_INT(nStation)];
IF pSt = 0 THEN
    sMsg := 'Station not ready yet, retry';
    RETURN;
END_IF
M_StartStation := pSt^.M_RequestStart(sMsg => sMsg);
END_METHOD

// RPC：停止所有 mover、中止站動作與自動循環。不受 ready / 模式限制，永遠接受。
{attribute 'TcRpcEnable'}
METHOD PUBLIC M_Stop : BOOL
VAR_OUTPUT
    sMsg : STRING;
END_VAR
bReqStop := TRUE;
IF bReady THEN
    sMsg := 'Stop accepted';
ELSE
    sMsg := 'Stop accepted (XTS not ready, movers may be unpowered)';
END_IF
M_Stop := TRUE;
END_METHOD

END_FUNCTION_BLOCK

// ---- POUs/FB_Mover.TcPOU
// 一個 XTS mover：MC_Power + CA 移動 / 停止 + 工件狀態。命令由 method 設旗標，body 每 cycle 執行。
// 前置：FB_XTS_Control 每 cycle 呼叫並寫入 stPermit；CA group 已 enable 才能移動。
FUNCTION_BLOCK FB_Mover
VAR_INPUT
    nIndex : INT;                   // mover 編號 1..cMoverCount
    stPermit : ST_CmdPermit;        // 總控每 cycle 寫入
    bPowerEnable : BOOL;            // 總控送電
    bResetCmd : BOOL;               // 總控初始化時的 reset
END_VAR
VAR_IN_OUT
    stAxis : AXIS_REF;
END_VAR
VAR_OUTPUT
    fPositionMm : LREAL;            // 環上位置 (mm), 0~cTrackLengthMm
    fVelocityMmS : LREAL;           // 實際速度 (mm/s)
    bPowered : BOOL;
    bBusy : BOOL;                   // 移動或停止中 (CA 排隊時也是 TRUE)
    bDone : BOOL;                   // 最後一次移動到位
    bError : BOOL;
    nErrorId : UDINT;
    bHasPart : BOOL;                // 有工件
    bPressed : BOOL;                // 已下壓
END_VAR
VAR
    fbPower : MC_Power;
    fbReset : MC_Reset;
    fbMove : Tc3_McCollisionAvoidance.MC_MoveAbsoluteCA;
    fbHalt : Tc3_McCollisionAvoidance.MC_HaltCA;
    fbMoveTimer : TON;
    eMoveState : E_MoveState;
    fTargetAbsMm : LREAL;           // NC 絕對目標 (mm)
    fCmdVelocityMmS : LREAL;        // 本次移動速度 (mm/s)
    bReqMove : BOOL;                // method 設，body 取走
    fReqPositionMm : LREAL;
    fReqVelocityMmS : LREAL;
    bReqStop : BOOL;
    bReqReset : BOOL;
    bResetBusy : BOOL;              // MC_Reset 執行中
END_VAR

stAxis.ReadStatus();
fbPower(Axis := stAxis, Enable := bPowerEnable, Enable_Positive := bPowerEnable,
    Enable_Negative := bPowerEnable, Override := 100);
bPowered := fbPower.Status;

// 命令只在這裡取走；method 只設 bReq*
IF bReqReset OR bResetCmd THEN
    bReqReset := FALSE;
    bResetBusy := TRUE;
END_IF
IF bReqStop THEN
    bReqStop := FALSE;
    bReqMove := FALSE;
    eMoveState := E_MoveState.StartHalt;
ELSIF bReqMove THEN
    bReqMove := FALSE;
    // 只往正方向走：目標 = 目前 + 環上差距
    fTargetAbsMm := stAxis.NcToPlc.ActPos + F_RingPosition(
        fPositionMm := fReqPositionMm - F_RingPosition(fPositionMm := stAxis.NcToPlc.ActPos, fLengthMm := GVL_Param.cTrackLengthMm),
        fLengthMm := GVL_Param.cTrackLengthMm);
    fCmdVelocityMmS := fReqVelocityMmS;
    bDone := FALSE;
    eMoveState := E_MoveState.StartMove;
END_IF

// MC FB 用上個 cycle 的狀態呼叫，StartMove / StartHalt 那個 cycle Execute = FALSE
fbReset(Axis := stAxis, Execute := bResetBusy);
fbMove(Axis := stAxis, Execute := (eMoveState = E_MoveState.Moving), Position := fTargetAbsMm,
    Velocity := fCmdVelocityMmS, Acceleration := GVL_Param.cMoverAccMmS2,
    Deceleration := GVL_Param.cMoverAccMmS2, Jerk := GVL_Param.cMoverJerkMmS3, Gap := GVL_Param.cCaGapMm);
fbHalt(Axis := stAxis, Execute := (eMoveState = E_MoveState.Halting), Deceleration := GVL_Param.cMoverAccMmS2,
    Jerk := GVL_Param.cMoverJerkMmS3, Gap := GVL_Param.cCaGapMm);
fbMoveTimer(IN := (eMoveState = E_MoveState.Moving), PT := GVL_Param.cMoveTimeout);

IF fbReset.Done OR fbReset.Error THEN
    bResetBusy := FALSE;
    IF fbReset.Done THEN
        bError := FALSE;
        nErrorId := 0;
    END_IF
END_IF

CASE eMoveState OF
E_MoveState.Idle:
    ;
E_MoveState.StartMove:
    eMoveState := E_MoveState.Moving;
E_MoveState.Moving:
    IF fbMove.Done THEN
        bDone := TRUE;
        eMoveState := E_MoveState.Idle;
    ELSIF fbMove.Error OR NOT bPowered THEN
        eMoveState := E_MoveState.Idle;
    ELSIF fbMoveTimer.Q THEN
        bError := TRUE;
        nErrorId := GVL_ErrorId.cErrMoveTimeout;
        eMoveState := E_MoveState.Idle;
    END_IF
E_MoveState.StartHalt:
    eMoveState := E_MoveState.Halting;
E_MoveState.Halting:
    IF fbHalt.Done OR fbHalt.Error OR NOT bPowered THEN
        eMoveState := E_MoveState.Idle;
    END_IF
ELSE
    bError := TRUE;
    nErrorId := GVL_ErrorId.cErrInvalidState;
    eMoveState := E_MoveState.Idle;
END_CASE

IF fbPower.Error THEN
    bError := TRUE;
    nErrorId := fbPower.ErrorID;
ELSIF fbMove.Error THEN
    bError := TRUE;
    nErrorId := fbMove.ErrorId;
ELSIF fbHalt.Error THEN
    bError := TRUE;
    nErrorId := fbHalt.ErrorId;
ELSIF stAxis.Status.Error THEN
    bError := TRUE;
    nErrorId := stAxis.Status.ErrorID;
END_IF

fPositionMm := F_RingPosition(fPositionMm := stAxis.NcToPlc.ActPos, fLengthMm := GVL_Param.cTrackLengthMm);
fVelocityMmS := stAxis.NcToPlc.ActVelo;
bBusy := (eMoveState <> E_MoveState.Idle);

// RPC：移到環上位置。需 ready + Manual。回 TRUE = 已接受 (不是已到位)。
{attribute 'TcRpcEnable'}
METHOD PUBLIC M_MoveTo : BOOL
VAR_INPUT
    fPosition : LREAL;      // 目標環上位置 (mm), 0 <= p < cTrackLengthMm
    fVelocity : LREAL;      // 速度 (mm/s), 0 < v <= cMaxVelocityMmS
END_VAR
VAR_OUTPUT
    sMsg : STRING;          // 拒絕原因或 'Accepted'
END_VAR
IF NOT F_CheckCmdAllowed(stPermit := stPermit, bNeedManual := TRUE, bNeedAuto := FALSE, sMsg => sMsg) THEN
    M_MoveTo := FALSE;
    RETURN;
END_IF
M_MoveTo := M_RequestMove(fPosition := fPosition, fVelocity := fVelocity, sMsg => sMsg);
END_METHOD

// 內部用 (總控與 M_MoveTo 共用)：檢查參數後設移動命令，不檢查模式
METHOD PUBLIC M_RequestMove : BOOL
VAR_INPUT
    fPosition : LREAL;      // 目標環上位置 (mm)
    fVelocity : LREAL;      // 速度 (mm/s)
END_VAR
VAR_OUTPUT
    sMsg : STRING;
END_VAR
M_RequestMove := FALSE;
IF bReqMove OR bReqStop THEN
    sMsg := 'Previous command not yet taken by PLC, retry';
ELSIF bError THEN
    sMsg := 'Mover in error, call M_InitialXTS';
ELSIF NOT bPowered THEN
    sMsg := 'Mover not powered';
ELSIF (fPosition < 0.0) OR (fPosition >= GVL_Param.cTrackLengthMm) THEN
    sMsg := CONCAT('Position out of range, 0 <= fPosition < ', LREAL_TO_STRING(GVL_Param.cTrackLengthMm));
ELSIF (fVelocity <= 0.0) OR (fVelocity > GVL_Param.cMaxVelocityMmS) THEN
    sMsg := CONCAT('Velocity out of range, 0 < fVelocity <= ', LREAL_TO_STRING(GVL_Param.cMaxVelocityMmS));
ELSE
    fReqPositionMm := fPosition;
    fReqVelocityMmS := fVelocity;
    bReqMove := TRUE;               // 旗標最後設
    sMsg := 'Accepted';
    M_RequestMove := TRUE;
END_IF
END_METHOD

// RPC：停止 (MC_HaltCA)。不受 ready / 模式限制，永遠接受。
{attribute 'TcRpcEnable'}
METHOD PUBLIC M_Stop : BOOL
VAR_OUTPUT
    sMsg : STRING;
END_VAR
bReqStop := TRUE;
IF bPowered THEN
    sMsg := 'Stop accepted';
ELSE
    sMsg := 'Not powered, nothing to stop';
END_IF
M_Stop := TRUE;
END_METHOD

// RPC：MC_Reset。需 ready + Manual；掉出 ready 後的復歸請用 M_InitialXTS。
{attribute 'TcRpcEnable'}
METHOD PUBLIC M_Reset : BOOL
VAR_OUTPUT
    sMsg : STRING;
END_VAR
IF NOT F_CheckCmdAllowed(stPermit := stPermit, bNeedManual := TRUE, bNeedAuto := FALSE, sMsg => sMsg) THEN
    M_Reset := FALSE;
    RETURN;
END_IF
bReqReset := TRUE;
sMsg := 'Reset accepted';
M_Reset := TRUE;
END_METHOD

// RPC：讀狀態，隨時可讀
{attribute 'TcRpcEnable'}
METHOD PUBLIC M_GetStatus : BOOL
VAR_OUTPUT
    fPosition : LREAL;      // 環上位置 (mm)
    fVelocity : LREAL;      // 實際速度 (mm/s)
    bBusy : BOOL;
    bError : BOOL;
    nErrorId : UDINT;
    bHasPart : BOOL;
    bPressed : BOOL;
    bPowered : BOOL;
END_VAR
fPosition := THIS^.fPositionMm;
fVelocity := THIS^.fVelocityMmS;
bBusy := THIS^.bBusy;
bError := THIS^.bError;
nErrorId := THIS^.nErrorId;
bHasPart := THIS^.bHasPart;
bPressed := THIS^.bPressed;
bPowered := THIS^.bPowered;
M_GetStatus := TRUE;
END_METHOD

// 內部用：站完成後由總控更新工件狀態
METHOD PUBLIC M_SetPart
VAR_INPUT
    bPart : BOOL;           // 有工件
    bPress : BOOL;          // 已下壓
END_VAR
bHasPart := bPart;
bPressed := bPress;
END_METHOD

END_FUNCTION_BLOCK

// ---- POUs/F_RingPosition.TcPOU
// 把位置換算到環上 0 ~ fLengthMm
FUNCTION F_RingPosition : LREAL
VAR_INPUT
    fPositionMm : LREAL;    // 任意位置 (mm)
    fLengthMm : LREAL;      // 環長 (mm), > 0
END_VAR

IF fLengthMm <= 0.0 THEN
    F_RingPosition := 0.0;
    RETURN;
END_IF
// TRUNC 回 DINT；|位置| 在 DINT 範圍內 (±2.1e9 mm) 不會溢位
F_RingPosition := fPositionMm - DINT_TO_LREAL(TRUNC(fPositionMm / fLengthMm)) * fLengthMm;
IF F_RingPosition < 0.0 THEN
    F_RingPosition := F_RingPosition + fLengthMm;
END_IF

END_FUNCTION

// ---- POUs/F_CheckCmdAllowed.TcPOU
// 命令允許檢查，所有 RPC 命令 method 都只呼叫這一個 (ready 閘門 + 模式鎖)
FUNCTION F_CheckCmdAllowed : BOOL
VAR_INPUT
    stPermit : ST_CmdPermit;
    bNeedManual : BOOL;     // 直接對 mover / 站的命令
    bNeedAuto : BOOL;       // 整線自動命令
END_VAR
VAR_OUTPUT
    sMsg : STRING;          // 拒絕原因，允許時為空字串
END_VAR

F_CheckCmdAllowed := FALSE;
IF NOT stPermit.bReady THEN
    sMsg := 'XTS not ready, call M_InitialXTS first';
ELSIF bNeedManual AND (stPermit.eMode <> E_XtsMode.Manual) THEN
    sMsg := 'Rejected in Auto mode, call M_SetMode(0) first';
ELSIF bNeedAuto AND (stPermit.eMode <> E_XtsMode.Auto) THEN
    sMsg := 'Needs Auto mode, call M_SetMode(1) first';
ELSE
    sMsg := '';
    F_CheckCmdAllowed := TRUE;
END_IF

END_FUNCTION

// ---- POUs/FB_StationLoad.TcPOU
// 第 1 站 Load：XYZ 從取料點夾工件放到 mover 上。mover 必須沒有工件。
FUNCTION_BLOCK FB_StationLoad EXTENDS FB_StationGantry

fPickXMm := GVL_Param.cGantryFeederXMm;
fPickYMm := GVL_Param.cGantryFeederYMm;
fPlaceXMm := GVL_Param.cGantryMoverXMm;
fPlaceYMm := GVL_Param.cGantryMoverYMm;
SUPER^(aAxis := aAxis);

METHOD PROTECTED M_CheckStart : BOOL
VAR_OUTPUT
    sMsg : STRING;
END_VAR
IF bMoverHasPart THEN
    sMsg := 'Mover already has a part';
    M_CheckStart := FALSE;
ELSE
    sMsg := '';
    M_CheckStart := TRUE;
END_IF
END_METHOD

END_FUNCTION_BLOCK

// ---- POUs/FB_StationGantry.TcPOU
// XYZ 取放站共用 (Load / Unload)：從 fPick 取料放到 fPlace。取放點由子類別 body 設定。
// 步驟：10 XY 到取料點 → 20 Z 下 → 30 夾 → 40 Z 上 → 50 XY 到放料點 → 60 Z 下 → 70 放 → 80 Z 上
FUNCTION_BLOCK FB_StationGantry EXTENDS FB_Station
VAR_IN_OUT
    aAxis : ARRAY[1..GVL_Param.cGantryAxisCount] OF AXIS_REF;     // X / Y / Z
END_VAR
VAR
    aSimAxis : ARRAY[1..GVL_Param.cGantryAxisCount] OF FB_SimAxis;
    aTargetMm : ARRAY[1..GVL_Param.cGantryAxisCount] OF LREAL;    // 本步目標 (mm)
    fPickXMm : LREAL;               // 取料點 X (mm)
    fPickYMm : LREAL;               // 取料點 Y (mm)
    fPlaceXMm : LREAL;              // 放料點 X (mm)
    fPlaceYMm : LREAL;              // 放料點 Y (mm)
    fbGripTimer : TON;
    bAxesHalt : BOOL;
    i : INT;
END_VAR

SUPER^();
fbGripTimer(IN := (nStep = 30) OR (nStep = 70), PT := GVL_Param.cGripTime);
// 奇數步 Execute = TRUE；偶數步先設目標、Execute = FALSE，產生下一個上升沿
bAxesPowered := TRUE;
bAxisError := FALSE;
FOR i := 1 TO GVL_Param.cGantryAxisCount DO
    aSimAxis[i](bPower := bPowerEnable,
        bExecute := (eState = E_StationState.Busy) AND ((nStep MOD 2) = 1),
        bHalt := bAxesHalt, bReset := bResetCmd, fTargetMm := aTargetMm[i],
        fVelocityMmS := GVL_Param.cGantryVelocityMmS, fAccMmS2 := GVL_Param.cGantryAccMmS2,
        stAxis := aAxis[i]);
    bAxesPowered := bAxesPowered AND aSimAxis[i].bPowered;
    bAxisError := bAxisError OR aSimAxis[i].bError;
END_FOR
fAxis1Mm := aSimAxis[GVL_Param.cAxisX].fActPosMm;
fAxis2Mm := aSimAxis[GVL_Param.cAxisY].fActPosMm;
fAxis3Mm := aSimAxis[GVL_Param.cAxisZ].fActPosMm;

METHOD PROTECTED M_Sequence
IF bAxisError THEN
    bSeqError := TRUE;
    FOR i := 1 TO GVL_Param.cGantryAxisCount DO
        IF aSimAxis[i].bError THEN
            nSeqErrorId := aSimAxis[i].nErrorId;
        END_IF
    END_FOR
    RETURN;
END_IF
CASE nStep OF
10:
    bAxesHalt := FALSE;
    M_SetTarget(fXMm := fPickXMm, fYMm := fPickYMm, fZMm := GVL_Param.cGantryZUpMm);
    nStep := 11;
11:
    IF M_AxesDone() THEN nStep := 20; END_IF
20:
    M_SetTarget(fXMm := fPickXMm, fYMm := fPickYMm, fZMm := GVL_Param.cGantryZDownMm);
    nStep := 21;
21:
    IF M_AxesDone() THEN nStep := 30; END_IF
30:
    bGripClosed := TRUE;
    IF fbGripTimer.Q THEN nStep := 40; END_IF
40:
    M_SetTarget(fXMm := fPickXMm, fYMm := fPickYMm, fZMm := GVL_Param.cGantryZUpMm);
    nStep := 41;
41:
    IF M_AxesDone() THEN nStep := 50; END_IF
50:
    M_SetTarget(fXMm := fPlaceXMm, fYMm := fPlaceYMm, fZMm := GVL_Param.cGantryZUpMm);
    nStep := 51;
51:
    IF M_AxesDone() THEN nStep := 60; END_IF
60:
    M_SetTarget(fXMm := fPlaceXMm, fYMm := fPlaceYMm, fZMm := GVL_Param.cGantryZDownMm);
    nStep := 61;
61:
    IF M_AxesDone() THEN nStep := 70; END_IF
70:
    bGripClosed := FALSE;
    IF fbGripTimer.Q THEN nStep := 80; END_IF
80:
    M_SetTarget(fXMm := fPlaceXMm, fYMm := fPlaceYMm, fZMm := GVL_Param.cGantryZUpMm);
    nStep := 81;
81:
    IF M_AxesDone() THEN bSeqDone := TRUE; END_IF
ELSE
    bSeqError := TRUE;
    nSeqErrorId := GVL_ErrorId.cErrInvalidState;
END_CASE
END_METHOD

METHOD PROTECTED M_Abort
bAxesHalt := TRUE;      // 夾爪狀態保留，工件可能還在夾爪上
END_METHOD

METHOD PRIVATE M_SetTarget
VAR_INPUT
    fXMm : LREAL;
    fYMm : LREAL;
    fZMm : LREAL;
END_VAR
aTargetMm[GVL_Param.cAxisX] := fXMm;
aTargetMm[GVL_Param.cAxisY] := fYMm;
aTargetMm[GVL_Param.cAxisZ] := fZMm;
END_METHOD

METHOD PRIVATE M_AxesDone : BOOL
VAR
    k : INT;
END_VAR
M_AxesDone := TRUE;
FOR k := 1 TO GVL_Param.cGantryAxisCount DO
    M_AxesDone := M_AxesDone AND aSimAxis[k].bDone;
END_FOR
END_METHOD

END_FUNCTION_BLOCK

// ---- POUs/FB_Station.TcPOU
// 站的共用底層：站狀態、占用、放行、步驟逾時。動作步驟由子類別覆寫 M_Sequence。
// 前置：FB_XTS_Control 每 cycle 寫入 stPermit、nMoverAtStation、bMoverHasPart、bMoverPressed 並呼叫。
FUNCTION_BLOCK FB_Station
VAR_INPUT
    nIndex : INT;                   // 站號 1..cStationCount
    stPermit : ST_CmdPermit;        // 總控每 cycle 寫入
    nMoverAtStation : INT;          // 停在站上的 mover，0 = 無
    bMoverHasPart : BOOL;           // 站上 mover 有工件
    bMoverPressed : BOOL;           // 站上 mover 已下壓
    bPowerEnable : BOOL;            // 站上軸送電
    bResetCmd : BOOL;               // 總控初始化時的 reset
    bAbort : BOOL;                  // 總控 Stop：中止動作、停軸
END_VAR
VAR_OUTPUT
    eState : E_StationState;
    nStep : INT;                    // 站內步驟，0 = 不在動作
    bOccupied : BOOL;               // 站內有 mover 或站在動作
    nMover : INT;                   // 處理中的 mover，0 = 無
    bBusy : BOOL;
    bDone : BOOL;
    bError : BOOL;
    nErrorId : UDINT;
    nDoneCount : UDINT;             // 完成次數
    bAxesPowered : BOOL;            // 站上軸全部送電
    bAxisError : BOOL;              // 站上軸 error，總控會因此掉出 ready
    fAxis1Mm : LREAL;               // X (mm)
    fAxis2Mm : LREAL;               // Y (mm)
    fAxis3Mm : LREAL;               // Z (mm)，往下為正
    bGripClosed : BOOL;             // 夾爪閉合
END_VAR
VAR
    bReqStart : BOOL;               // method 設，body 取走
    bReqRelease : BOOL;
    bReqReset : BOOL;
    fbStepTimer : TON;
    nStepLast : INT;
    bSeqDone : BOOL;                // M_Sequence 回報
    bSeqError : BOOL;
    nSeqErrorId : UDINT;
END_VAR

fbStepTimer(IN := (eState = E_StationState.Busy) AND (nStep = nStepLast), PT := GVL_Param.cStationStepTimeout);
nStepLast := nStep;

IF bResetCmd OR bReqReset THEN
    bReqReset := FALSE;
    IF eState = E_StationState.Busy THEN
        M_Abort();
    END_IF
    IF eState <> E_StationState.Done THEN
        eState := E_StationState.Idle;
        nStep := 0;
        nMover := 0;
    END_IF
    nErrorId := 0;
END_IF
IF bAbort AND (eState = E_StationState.Busy) THEN
    M_Abort();
    eState := E_StationState.Idle;
    nStep := 0;
    nMover := 0;
END_IF

CASE eState OF
E_StationState.Idle:
    IF bReqStart THEN
        nMover := nMoverAtStation;
        nStep := 10;
        eState := E_StationState.Busy;
    END_IF
E_StationState.Busy:
    bSeqDone := FALSE;
    bSeqError := FALSE;
    M_Sequence();
    IF bSeqError THEN
        nErrorId := nSeqErrorId;
        eState := E_StationState.Error;
    ELSIF bSeqDone THEN
        nDoneCount := nDoneCount + 1;
        nStep := 0;
        eState := E_StationState.Done;
    ELSIF fbStepTimer.Q THEN
        M_Abort();
        nErrorId := GVL_ErrorId.cErrStationTimeout;
        eState := E_StationState.Error;
    END_IF
E_StationState.Done:
    IF bReqRelease THEN
        nMover := 0;
        eState := E_StationState.Idle;
    END_IF
E_StationState.Error:
    ;
ELSE
    nErrorId := GVL_ErrorId.cErrInvalidState;
    eState := E_StationState.Error;
END_CASE
// 沒在對應狀態被取走的請求直接丟掉
bReqStart := FALSE;
bReqRelease := FALSE;

bBusy := (eState = E_StationState.Busy);
bDone := (eState = E_StationState.Done);
bError := (eState = E_StationState.Error);
bOccupied := (nMoverAtStation <> 0) OR (eState <> E_StationState.Idle);

// RPC：手動跑一次站動作。需 ready + Manual、站 Idle、站上有 mover。
{attribute 'TcRpcEnable'}
METHOD PUBLIC M_Start : BOOL
VAR_OUTPUT
    sMsg : STRING;
END_VAR
IF NOT F_CheckCmdAllowed(stPermit := stPermit, bNeedManual := TRUE, bNeedAuto := FALSE, sMsg => sMsg) THEN
    M_Start := FALSE;
    RETURN;
END_IF
M_Start := M_RequestStart(sMsg => sMsg);
END_METHOD

// 內部用 (總控自動循環與 M_Start 共用)：檢查站狀態後設啟動命令，不檢查模式
METHOD PUBLIC M_RequestStart : BOOL
VAR_OUTPUT
    sMsg : STRING;
END_VAR
M_RequestStart := FALSE;
IF bReqStart THEN
    sMsg := 'Previous command not yet taken by PLC, retry';
ELSIF eState <> E_StationState.Idle THEN
    sMsg := 'Station not idle (busy, waiting release or error)';
ELSIF nMoverAtStation = 0 THEN
    sMsg := 'No mover at station';
ELSIF M_CheckStart(sMsg => sMsg) THEN
    bReqStart := TRUE;
    sMsg := 'Accepted';
    M_RequestStart := TRUE;
END_IF
END_METHOD

// RPC：放行 (Done -> Idle)。需 ready + Manual。
{attribute 'TcRpcEnable'}
METHOD PUBLIC M_Release : BOOL
VAR_OUTPUT
    sMsg : STRING;
END_VAR
IF NOT F_CheckCmdAllowed(stPermit := stPermit, bNeedManual := TRUE, bNeedAuto := FALSE, sMsg => sMsg) THEN
    M_Release := FALSE;
    RETURN;
END_IF
M_Release := M_RequestRelease(sMsg => sMsg);
END_METHOD

// 內部用：站在 Done 才放行
METHOD PUBLIC M_RequestRelease : BOOL
VAR_OUTPUT
    sMsg : STRING;
END_VAR
IF eState = E_StationState.Done THEN
    bReqRelease := TRUE;
    sMsg := 'Accepted';
    M_RequestRelease := TRUE;
ELSE
    sMsg := 'Station not in Done, nothing to release';
    M_RequestRelease := FALSE;
END_IF
END_METHOD

// RPC：清站的 Error 回 Idle (站上軸 MC_Reset 走 M_InitialXTS)。需 ready + Manual。
{attribute 'TcRpcEnable'}
METHOD PUBLIC M_Reset : BOOL
VAR_OUTPUT
    sMsg : STRING;
END_VAR
IF NOT F_CheckCmdAllowed(stPermit := stPermit, bNeedManual := TRUE, bNeedAuto := FALSE, sMsg => sMsg) THEN
    M_Reset := FALSE;
    RETURN;
END_IF
bReqReset := TRUE;
sMsg := 'Reset accepted';
M_Reset := TRUE;
END_METHOD

// RPC：讀狀態，隨時可讀
{attribute 'TcRpcEnable'}
METHOD PUBLIC M_GetStatus : BOOL
VAR_OUTPUT
    nState : INT;           // E_StationState 值
    nStepNow : INT;
    bOccupiedNow : BOOL;
    nMoverNow : INT;
    bErrorNow : BOOL;
    nErrorIdNow : UDINT;
    nDone : UDINT;
    fAxisX : LREAL;         // (mm)
    fAxisY : LREAL;         // (mm)
    fAxisZ : LREAL;         // (mm)
END_VAR
CASE eState OF
E_StationState.Idle:  nState := 0;
E_StationState.Busy:  nState := 10;
E_StationState.Done:  nState := 20;
E_StationState.Error: nState := 900;
ELSE
    nState := -1;
END_CASE
nStepNow := nStep;
bOccupiedNow := bOccupied;
nMoverNow := nMover;
bErrorNow := bError;
nErrorIdNow := nErrorId;
nDone := nDoneCount;
fAxisX := fAxis1Mm;
fAxisY := fAxis2Mm;
fAxisZ := fAxis3Mm;
M_GetStatus := TRUE;
END_METHOD

// 內部用：給總控組 ST_LineStatus
METHOD PUBLIC M_GetStatusStruct : ST_StationStatus
M_GetStatusStruct.eState := eState;
M_GetStatusStruct.nStep := nStep;
M_GetStatusStruct.bOccupied := bOccupied;
M_GetStatusStruct.nMover := nMover;
M_GetStatusStruct.bError := bError;
M_GetStatusStruct.nErrorId := nErrorId;
M_GetStatusStruct.nDoneCount := nDoneCount;
M_GetStatusStruct.fAxis1Mm := fAxis1Mm;
M_GetStatusStruct.fAxis2Mm := fAxis2Mm;
M_GetStatusStruct.fAxis3Mm := fAxis3Mm;
M_GetStatusStruct.bGripClosed := bGripClosed;
END_METHOD

// 子類別覆寫：檢查站上 mover 的工件狀態可否開始
METHOD PROTECTED M_CheckStart : BOOL
VAR_OUTPUT
    sMsg : STRING;
END_VAR
sMsg := '';
M_CheckStart := TRUE;
END_METHOD

// 子類別覆寫：每 cycle 推進一步，完成設 bSeqDone，失敗設 bSeqError / nSeqErrorId
METHOD PROTECTED M_Sequence
bSeqDone := TRUE;
END_METHOD

// 子類別覆寫：中止時停軸
METHOD PROTECTED M_Abort
;
END_METHOD

END_FUNCTION_BLOCK

// ---- POUs/FB_SimAxis.TcPOU
// 單一 NC 模擬軸 (站上 XYZ / 下壓軸)：送電、絕對移動、停止、reset。每 cycle 呼叫。
FUNCTION_BLOCK FB_SimAxis
VAR_INPUT
    bPower : BOOL;
    bExecute : BOOL;            // 上升沿移到 fTargetMm
    bHalt : BOOL;               // 上升沿停止，優先於 bExecute
    bReset : BOOL;              // 上升沿 MC_Reset，並清 bError
    fTargetMm : LREAL;          // 目標位置 (mm)
    fVelocityMmS : LREAL;       // 速度 (mm/s), > 0
    fAccMmS2 : LREAL;           // 加減速度 (mm/s2), > 0
END_VAR
VAR_IN_OUT
    stAxis : AXIS_REF;
END_VAR
VAR_OUTPUT
    bPowered : BOOL;
    bBusy : BOOL;
    bDone : BOOL;               // 本次移動到位，bExecute 回 FALSE 時清掉
    bError : BOOL;
    nErrorId : UDINT;
    fActPosMm : LREAL;          // 實際位置 (mm)
END_VAR
VAR
    fbPower : MC_Power;
    fbReset : MC_Reset;
    fbMove : MC_MoveAbsolute;
    fbHalt : MC_Halt;
END_VAR

stAxis.ReadStatus();
fbPower(Axis := stAxis, Enable := bPower, Enable_Positive := bPower, Enable_Negative := bPower, Override := 100);
fbReset(Axis := stAxis, Execute := bReset);
fbMove(Axis := stAxis, Execute := bExecute AND fbPower.Status AND NOT bHalt,
    Position := fTargetMm, Velocity := fVelocityMmS, Acceleration := fAccMmS2, Deceleration := fAccMmS2);
fbHalt(Axis := stAxis, Execute := bHalt AND fbPower.Status, Deceleration := fAccMmS2);
bPowered := fbPower.Status;
bBusy := fbMove.Busy OR fbHalt.Busy;
bDone := fbMove.Done;
fActPosMm := stAxis.NcToPlc.ActPos;
IF bReset THEN
    bError := FALSE;
    nErrorId := 0;
END_IF
IF fbPower.Error THEN
    bError := TRUE;
    nErrorId := fbPower.ErrorID;
ELSIF fbMove.Error THEN
    bError := TRUE;
    nErrorId := fbMove.ErrorID;
ELSIF fbHalt.Error THEN
    bError := TRUE;
    nErrorId := fbHalt.ErrorID;
ELSIF stAxis.Status.Error THEN
    bError := TRUE;
    nErrorId := stAxis.Status.ErrorID;
END_IF

END_FUNCTION_BLOCK

// ---- POUs/FB_StationPress.TcPOU
// 第 2 站 Press：下壓軸下降 → 保壓 → 上升。mover 必須有工件且還沒下壓。
// 步驟：10 下降 → 20 保壓 → 30 上升
FUNCTION_BLOCK FB_StationPress EXTENDS FB_Station
VAR_IN_OUT
    stAxis : AXIS_REF;              // 下壓軸 (Z)
END_VAR
VAR
    fbPressAxis : FB_SimAxis;
    fTargetMm : LREAL;              // 本步目標 (mm)
    fbHoldTimer : TON;
    bAxisHalt : BOOL;
END_VAR

SUPER^();
fbHoldTimer(IN := (nStep = 20), PT := GVL_Param.cPressHoldTime);
fbPressAxis(bPower := bPowerEnable,
    bExecute := (eState = E_StationState.Busy) AND ((nStep MOD 2) = 1),
    bHalt := bAxisHalt, bReset := bResetCmd, fTargetMm := fTargetMm,
    fVelocityMmS := GVL_Param.cGantryVelocityMmS, fAccMmS2 := GVL_Param.cGantryAccMmS2,
    stAxis := stAxis);
bAxesPowered := fbPressAxis.bPowered;
bAxisError := fbPressAxis.bError;
fAxis3Mm := fbPressAxis.fActPosMm;

METHOD PROTECTED M_CheckStart : BOOL
VAR_OUTPUT
    sMsg : STRING;
END_VAR
IF NOT bMoverHasPart THEN
    sMsg := 'Mover has no part to press';
    M_CheckStart := FALSE;
ELSIF bMoverPressed THEN
    sMsg := 'Part already pressed';
    M_CheckStart := FALSE;
ELSE
    sMsg := '';
    M_CheckStart := TRUE;
END_IF
END_METHOD

METHOD PROTECTED M_Sequence
IF bAxisError THEN
    bSeqError := TRUE;
    nSeqErrorId := fbPressAxis.nErrorId;
    RETURN;
END_IF
CASE nStep OF
10:
    bAxisHalt := FALSE;
    fTargetMm := GVL_Param.cPressZDownMm;
    nStep := 11;
11:
    IF fbPressAxis.bDone THEN nStep := 20; END_IF
20:
    IF fbHoldTimer.Q THEN nStep := 30; END_IF
30:
    fTargetMm := GVL_Param.cGantryZUpMm;
    nStep := 31;
31:
    IF fbPressAxis.bDone THEN bSeqDone := TRUE; END_IF
ELSE
    bSeqError := TRUE;
    nSeqErrorId := GVL_ErrorId.cErrInvalidState;
END_CASE
END_METHOD

METHOD PROTECTED M_Abort
bAxisHalt := TRUE;
END_METHOD

END_FUNCTION_BLOCK

// ---- POUs/FB_StationUnload.TcPOU
// 第 3 站 Unload：XYZ 從 mover 夾走工件放到出料點。mover 必須有工件。
FUNCTION_BLOCK FB_StationUnload EXTENDS FB_StationGantry

fPickXMm := GVL_Param.cGantryMoverXMm;
fPickYMm := GVL_Param.cGantryMoverYMm;
fPlaceXMm := GVL_Param.cGantryOutXMm;
fPlaceYMm := GVL_Param.cGantryOutYMm;
SUPER^(aAxis := aAxis);

METHOD PROTECTED M_CheckStart : BOOL
VAR_OUTPUT
    sMsg : STRING;
END_VAR
IF NOT bMoverHasPart THEN
    sMsg := 'Mover has no part to unload';
    M_CheckStart := FALSE;
ELSE
    sMsg := '';
    M_CheckStart := TRUE;
END_IF
END_METHOD

END_FUNCTION_BLOCK

// ---- POUs/FB_CaGroup.TcPOU
// CA group 管理：mover 加進 group、enable；bEnable 回 FALSE 時 disable 並 ungroup。
FUNCTION_BLOCK FB_CaGroup
VAR_INPUT
    bEnable : BOOL;
    bReset : BOOL;
END_VAR
VAR_IN_OUT
    Group : Tc3_McCoordinatedMotion.AXES_GROUP_REF;
    Axes : ARRAY[1..GVL_Param.cMoverCount] OF AXIS_REF;
END_VAR
VAR_OUTPUT
    bReady : BOOL;          // group enable 完成且軸數正確
    bError : BOOL;
    nErrorId : UDINT;
    nState : UINT;          // 0 idle, 10 add, 20 enable, 30 ready, 80 disable, 90 ungroup
    nAxesCount : UDINT;
END_VAR
VAR
    aAdd : ARRAY[1..GVL_Param.cMoverCount] OF Tc3_McCoordinatedMotion.MC_AddAxisToGroup;
    fbEnable : Tc3_McCoordinatedMotion.MC_GroupEnable;
    fbDisable : Tc3_McCoordinatedMotion.MC_GroupDisable;
    fbUngroup : Tc3_McCoordinatedMotion.MC_UngroupAllAxes;
    fbReset : Tc3_McCoordinatedMotion.MC_GroupReset;
    bAllAdded : BOOL;
    i : INT;
END_VAR
VAR CONSTANT
    cErrNoGroup : UDINT := 16#E202;     // CA group 物件不存在 (GroupOID = 0)
END_VAR

// 逾時由 FB_XTS_Control 的初始化步驟計時 (cInitStepTimeout)
nAxesCount := Group.NcToPlc.Common.GroupAxesCount;
fbReset(AxesGroup := Group, Execute := bReset);
IF bReset THEN
    bError := FALSE;
    nErrorId := 0;
    nState := 0;
END_IF
IF NOT bEnable AND (nState > 0) AND (nState < 80) THEN
    nState := 80;
END_IF
bAllAdded := TRUE;
FOR i := 1 TO GVL_Param.cMoverCount DO
    aAdd[i](AxesGroup := Group, Axis := Axes[i], Execute := (nState = 10),
        IdentInGroup := Tc3_McCoordinatedMotion.UDINT_TO_IDENTINGROUP(INT_TO_UDINT(i)));
    bAllAdded := bAllAdded AND aAdd[i].Done;
    IF aAdd[i].Error THEN
        bError := TRUE;
        nErrorId := aAdd[i].ErrorId;
    END_IF
END_FOR
fbEnable(AxesGroup := Group, Execute := (nState = 20));
fbDisable(AxesGroup := Group, Execute := (nState = 80));
fbUngroup(AxesGroup := Group, Execute := (nState = 90));
IF fbUngroup.Error THEN
    bError := TRUE;
    nErrorId := fbUngroup.ErrorId;
END_IF
IF fbEnable.Error THEN
    bError := TRUE;
    nErrorId := fbEnable.ErrorId;
END_IF
IF fbDisable.Error THEN
    bError := TRUE;
    nErrorId := fbDisable.ErrorId;
END_IF
CASE nState OF
0:
    IF bEnable AND NOT bError AND NOT bReset THEN
        IF Group.NcToPlc.Common.GroupOID = 0 THEN
            bError := TRUE;
            nErrorId := cErrNoGroup;
        ELSIF nAxesCount = INT_TO_UDINT(GVL_Param.cMoverCount) THEN
            nState := 20;
        ELSE
            nState := 10;
        END_IF
    END_IF
10:
    IF bAllAdded THEN
        nState := 20;
    END_IF
20:
    IF fbEnable.Done THEN
        nState := 30;
    END_IF
30:
    ;
80:
    IF fbDisable.Done AND (Group.NcToPlc.Common.GroupStatus.State =
        Tc3_McCoordinatedMotion.MC_GROUP_STATE.mcGroupStateDisabled) THEN
        nState := 90;
    END_IF
90:
    IF fbUngroup.Done AND (nAxesCount = 0) THEN
        nState := 0;
    END_IF
ELSE
    bError := TRUE;
    nErrorId := GVL_ErrorId.cErrInvalidState;
    nState := 0;
END_CASE
IF Group.NcToPlc.Common.GroupErrorId <> 0 THEN
    bError := TRUE;
    nErrorId := Group.NcToPlc.Common.GroupErrorId;
END_IF
bReady := (nState = 30) AND (nAxesCount = INT_TO_UDINT(GVL_Param.cMoverCount)) AND NOT bError;

END_FUNCTION_BLOCK

// ---- POUs/F_InitStepName.TcPOU
// 初始化步驟名稱，給 sInitMsg 用
FUNCTION F_InitStepName : STRING
VAR_INPUT
    eStep : E_InitStep;
END_VAR

CASE eStep OF
E_InitStep.Idle:            F_InitStepName := 'Idle';
E_InitStep.Reset:           F_InitStepName := 'Reset';
E_InitStep.InitEnvironment: F_InitStepName := 'InitEnvironment';
E_InitStep.WaitMovers:      F_InitStepName := 'WaitMovers';
E_InitStep.FindMover1:      F_InitStepName := 'FindMover1';
E_InitStep.FindMover1Wait:  F_InitStepName := 'FindMover1Wait';
E_InitStep.PowerOn:         F_InitStepName := 'PowerOn';
E_InitStep.EnableGroup:     F_InitStepName := 'EnableGroup';
E_InitStep.Ready:           F_InitStepName := 'Ready';
E_InitStep.Error:           F_InitStepName := 'Error';
ELSE
    F_InitStepName := 'Unknown';
END_CASE

END_FUNCTION
